// TIA Portal V21 export
// export: Created 2026-11-11T00:47:41.3931214Z, ExportSetting WithDefaults, DisplayName Totally Integrated Automation Portal, DisplayVersion V21 Update 3, DisplayName STEP 7 Professional, DisplayVersion V21 Update 3, DisplayName STEP 7 Safety, DisplayVersion V21, DisplayName Tech WebApplication, DisplayVersion V21, DisplayName WinCC Basic/Comfort/Advanced, DisplayVersion V21 Update 3, DisplayName WinCC Unified, DisplayVersion V21 Update 3
FUNCTION_BLOCK "FB_Fbd_ex156"   // FB164, FBD
{ S7_Optimized_Access := 'TRUE' }
VERSION : 0.1
// stored: AutoNumber true, IsIECCheckEnabled false, IsRetainMemResEnabled false, MemoryReserve 100, SetENOAutomatically false, UDAEnableTagReadback false
   VAR_INPUT
      v_laddr : HW_IO;
   END_VAR
   VAR_OUTPUT
      v_ret_val : Int;
      v_piaddr : UDInt;
      v_picount : UInt;
      v_pqaddr : UDInt;
      v_pqcount : UInt;
   END_VAR
BEGIN

REGION Network 1: RD_ADDR - Determine IO addresses from the hardware identifier
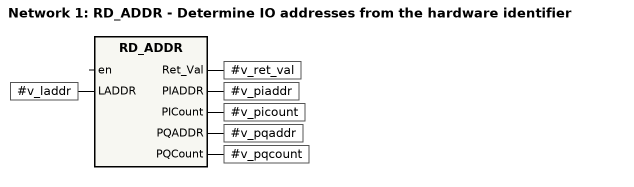
   #v_ret_val := RD_ADDR(LADDR := #v_laddr,
                         PIADDR => #v_piaddr,
                         PICount => #v_picount,
                         PQADDR => #v_pqaddr,
                         PQCount => #v_pqcount);
END_REGION
END_FUNCTION_BLOCK
